{attribute 'qualified_only'}
VAR_GLOBAL
	VTD:  VTD_Settings_DUT;
	ECnv:  ECnv_Settings_DUT;
	LCnv:  ARRAY[1..6] OF Buffer_Cnv_Settings_DUT;
	Turn_Table: Turn_Table_Settings_DUT;
	TBCnv:  TBCnv_Settings_DUT;
	Pop_Up_Cnv: ARRAY[1..2] OF PopUp_Settings_DUT;
	Roller_Cnv: ARRAY[1..5] OF Roller_Settings_DUT;
	Chain_Cnv: Chain_Settings_DUT;
// 	Shuttle_MQTT:  MQTT_Settings;
	System:  System_Settings_DUT;
END_VAR

(* stored: Version 1.1.0.1
   GVL Settings: Id {9b82498a-e9a0-4bb6-a6fe-ce7c787e0820} *)
